Fanuc KAREL source: kb00108.KL

PROGRAM KB00108
%STACKSIZE=65535
%PRIORITY=65535
%NOLOCKGROUP
VAR
P1 : INTEGER
P2 : INTEGER
P4 : ARRAY[4] OF INTEGER
P5 : INTEGER
-- UNRESOLVED DECLARATIONS (source type spelling not recovered)
-- P3 : TYPE_0x1100 (type_u16=0x1100)
BEGIN
P1=1
P2=1
P4[1]=1
P5=1
INSERT_QUEUE(P1,P2,P3,P4,P5)
END KB00108
